PROGRAM Parallel
  VAR
    TON0 : TON;
    h05_out : BOOL;
    CTU0 : CTU;
    h05_a : BOOL;
    h05_b : BOOL;
    h05_r : BOOL;
    h06_en : BOOL;
    h06_y1 : BOOL;
    h06_y2 : BOOL;
    h06_y3 : BOOL;
    h06_y4 : BOOL;
    TON1 : TON;
    h06_a1 : BOOL;
    TOF0 : TOF;
    h06_b1 : BOOL;
    CTU1 : CTU;
    h06_c1 : BOOL;
    h06_r : BOOL;
    h06_cv : INT;
    h09_out : BOOL;
    TON2 : TON;
    TOF1 : TOF;
    h09_a : BOOL;
    h09_b : BOOL;
    h09_c : BOOL;
    h09_d : BOOL;
  END_VAR

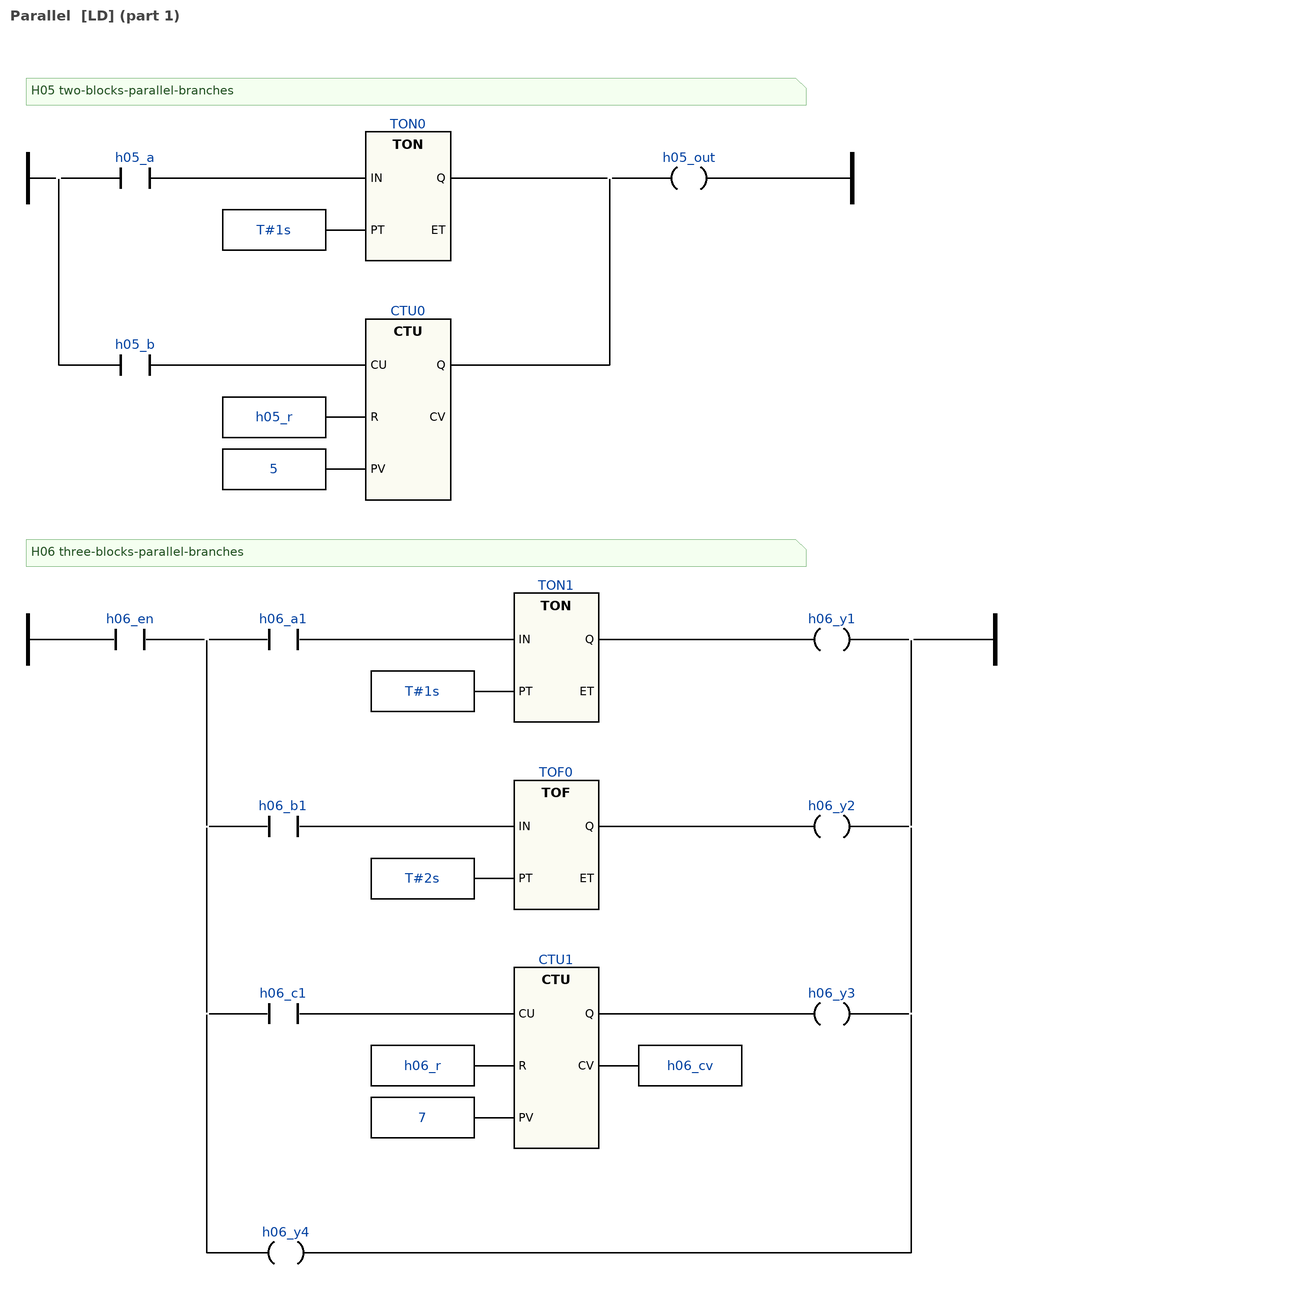
(* LD diagram, written out as Structured Text *)
(* H05 two-blocks-parallel-branches *)
TON0(IN := h05_a, PT := T#1s);
CTU0(CU := h05_b, R := h05_r, PV := 5);
h05_out := TON0.Q OR CTU0.Q;
(* H06 three-blocks-parallel-branches *)
TON1(IN := h06_en AND h06_a1, PT := T#1s);
h06_y1 := TON1.Q;
TOF0(IN := h06_en AND h06_b1, PT := T#2s);
h06_y2 := TOF0.Q;
CTU1(CU := h06_en AND h06_c1, R := h06_r, PV := 7);
h06_y3 := CTU1.Q;
h06_y4 := h06_en;
h06_cv := CTU1.CV;
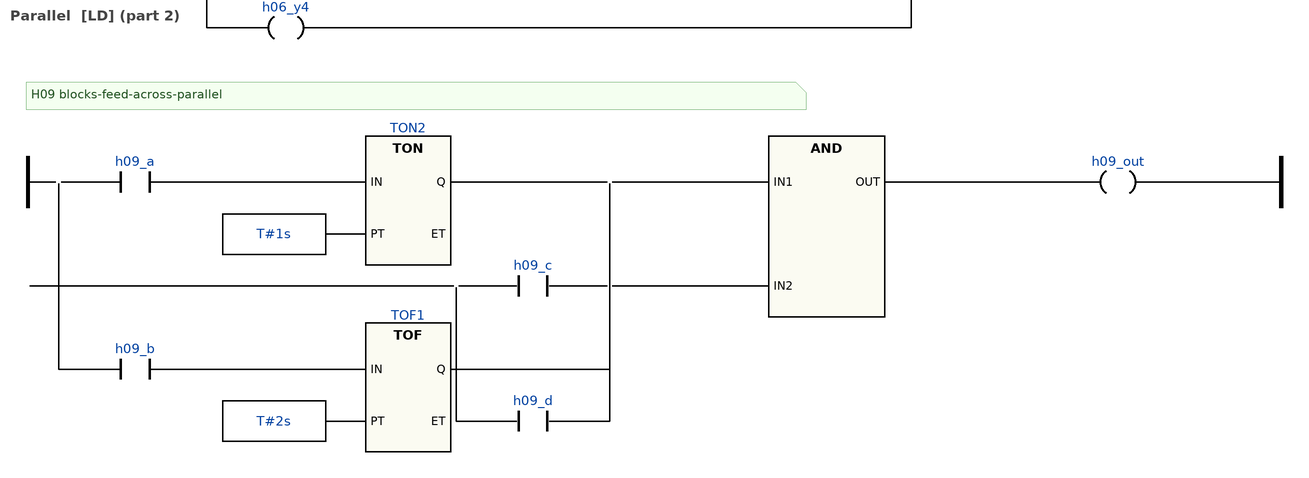
(* H09 blocks-feed-across-parallel *)
TON2(IN := h09_a, PT := T#1s);
TOF1(IN := h09_b, PT := T#2s);
h09_out := (TON2.Q OR TOF1.Q) AND (h09_c OR h09_d);
END_PROGRAM
